Fanuc KAREL source: KS00021.KL

PROGRAM KS00021
%NOLOCKGROUP
TYPE
  REC_T = STRUCTURE
    VALUE: INTEGER
    FLAG: BOOLEAN
  ENDSTRUCTURE
VAR
  A: FILE
  B: FILE
  FLAG: BOOLEAN
  N: INTEGER
  STATUS: INTEGER
  PN: STRING[80]
  VN: STRING[80]
BEGIN
  PN = ''
  VN = 'A'
  SET_VAR(N, PN, VN, A, STATUS)
END KS00021
